{attribute 'qualified_only'}
VAR_GLOBAL
	// global logger provider
	resource: FB_Resource(schemaUrl:='');
	loggerProvider: FB_LoggerProvider(resource:=resource);
	
	// global tracer provider
	sampler: FB_Sampler_AlwaysOn();
	idGenerator: FB_IdGenerator(nTraceIds:=5, nSpanIds:=5);
	tracerProvider: FB_TracerProvider(resource:=resource, idGenerator:=idGenerator, sampler:=sampler);

	// the master's interface over ADS: it writes command and reads status
	command: ST_SkidCommand;
	status: ST_SkidStatus;
END_VAR

(* stored: Version 1.1.0.1
   GVL GVL: Id {0fa68e8f-021a-4890-95b7-2639fe32abe1} *)
